(* IEC 61131-3 sources: plcassist-cli/packages/volt-lsp-iec/test-corpus/pro2193/Device/Plc Logic/Application/09 Misc/Library Manager/OMAC_PackML_State_Machine, 6 files *)

(* ---- GVL.gvl ---- *)
VAR_GLOBAL
	GC_USIMAXMODES : USINT := 10;
END_VAR

(* ---- IUNITMODE.itf ---- *)
INTERFACE IUNITMODE
END_INTERFACE

METHOD ABORT : BOOL
END_METHOD

METHOD ACTINGSTATECOMPLETED : BOOL
END_METHOD

METHOD CLEAR : BOOL
END_METHOD

METHOD HOLD : BOOL
END_METHOD

METHOD RESET : BOOL
END_METHOD

METHOD START : BOOL
END_METHOD

METHOD STOP : BOOL
END_METHOD

METHOD SUSPEND : BOOL
END_METHOD

METHOD UNHOLD : BOOL
END_METHOD

METHOD UNSUSPEND : BOOL
END_METHOD

METHOD ALLOWSENTERING : BOOL
VAR_INPUT
	E : State;
END_VAR
END_METHOD

METHOD ENTER : BOOL
VAR_INPUT
	E : State;
END_VAR
END_METHOD

METHOD NEXTSTATE : State
VAR_INPUT
	E : State;
END_VAR
END_METHOD

(* ---- GLOBALTEXTLIST.fb ---- *)
FUNCTION_BLOCK GLOBALTEXTLIST
VAR
	M_TEXTLISTFILE : STRING(255);
	_STNAMESPACE : STRING;
END_VAR
END_FUNCTION_BLOCK

(* ---- IMAGEPOOL.fb ---- *)
FUNCTION_BLOCK IMAGEPOOL
VAR
	M_STNAMESPACE : STRING(80);
	M_STHELPVARID : STRING;
	M_STHELPVARPATH : STRING(255);
	M_STHELP : STRING;
	M_REGISTERIMAGES : BOOL := TRUE;
END_VAR
END_FUNCTION_BLOCK

METHOD FB_INIT : BOOL
VAR_INPUT
	BINITRETAINS : BOOL;
	BINCOPYCODE : BOOL;
END_VAR
END_METHOD

METHOD FB_REINIT : BOOL
END_METHOD

METHOD FB_EXIT : BOOL
VAR_INPUT
	BINCOPYCODE : BOOL;
END_VAR
END_METHOD

(* ---- UNITMODE.fb ---- *)
FUNCTION_BLOCK UNITMODE
VAR_INPUT
	SNAME : STRING;
	DWSUPPORTEDSTATES : DWORD := 2#11111111111111111;
	DWALLOWSLEAVINGFROMSTATES : DWORD := (State.Stopped OR State.Aborted);
	DWALLOWSENTERINGINTOSTATES : DWORD := (State.Stopped OR State.Aborted);
	EINITIALSTATE : State;
	XACTIVE : BOOL;
END_VAR
VAR
	ESTATE : State := State.Invalid;
	BINIT : BOOL;
	ACTIVE : BOOL;
	ALLOWSLEAVING : BOOL;
	CURRENTSTATE : State;
	NAME : STRING;
	SUPPORTEDSTATES : DWORD;
END_VAR
END_FUNCTION_BLOCK

METHOD ABORT : BOOL
END_METHOD

METHOD ACTINGSTATECOMPLETED : BOOL
END_METHOD

METHOD CLEAR : BOOL
END_METHOD

METHOD HOLD : BOOL
END_METHOD

METHOD RESET : BOOL
END_METHOD

METHOD START : BOOL
END_METHOD

METHOD STOP : BOOL
END_METHOD

METHOD SUSPEND : BOOL
END_METHOD

METHOD UNHOLD : BOOL
END_METHOD

METHOD UNSUSPEND : BOOL
END_METHOD

METHOD ALLOWSENTERING : BOOL
VAR_INPUT
	E : State;
END_VAR
END_METHOD

METHOD ENTER : BOOL
VAR_INPUT
	E : State;
END_VAR
END_METHOD

METHOD NEXTSTATE : State
VAR_INPUT
	E : State;
END_VAR
END_METHOD

(* ---- UNITMODEMANAGER.fb ---- *)
FUNCTION_BLOCK UNITMODEMANAGER
VAR
	APUM : ARRAY [1..gc_usiMaxModes] OF IUnitMode;
	USINUMBEROFUMS : USINT := 0;
	USIACTUALUM : USINT;
	ACTIVEUNITMODE : IUnitMode;
	ACTIVEUNITMODENUMBER : USINT;
END_VAR
END_FUNCTION_BLOCK

METHOD ALLOWSSWITCHINGTO : BOOL
VAR_INPUT
	USI : USINT;
END_VAR
END_METHOD

METHOD FINDMODE : USINT
VAR_INPUT
	SNAME : STRING;
END_VAR
END_METHOD

METHOD REGISTER : BOOL
VAR_INPUT
	PUM : IUnitMode;
END_VAR
END_METHOD

METHOD SWITCHUNITMODE : BOOL
VAR_INPUT
	SNEWMODENAME : STRING;
END_VAR
END_METHOD
